(* PLC project boiler-plc210.project, CODESYS CODESYS V3.5 SP17 Patch 3 *)
(* stored: creationDateTime 2026-10-20T00:00:00, modificationDateTime 2026-10-20T00:00:00 *)
(* Синтетический экспорт: логика — corpus/boiler-plc210/src, слой ОВЕН — tools/corpus/owen_overlay.py (проба P7 не выполнялась) *)

// Назначение: состояние котла (вымышленная котельная №3, ПЛК210 — синтетический слой ОВЕН).
// Автор:      kr0nsch
// Версия:     0.1.0
// Документ:   corpus/boiler-plc210/README.md
{attribute 'qualified_only'}
TYPE E_BoilerState :
(
    Off := 0,       // остановлен
    Run := 1,       // работа
    Fault := 2      // авария горелки
) INT;
END_TYPE

// Назначение: отопительный график: уставка подачи по наружной температуре (линейно, с ограничением).
// Автор:      kr0nsch
// Версия:     0.1.0
// Документ:   corpus/boiler-plc210/README.md
FUNCTION F_HeatingCurve : REAL
VAR_INPUT
    rTOutdoor_C : REAL;     // наружная температура, °C
    rSpBase_C : REAL;       // уставка при 0 °C
END_VAR
VAR CONSTANT
    SLOPE : REAL := -1.2;   // наклон графика, °C/°C
    SP_MIN : REAL := 35.0;  // минимум подачи, °C
    SP_MAX : REAL := 95.0;  // максимум подачи, °C
END_VAR

            F_HeatingCurve := LIMIT(SP_MIN, rSpBase_C + SLOPE * rTOutdoor_C, SP_MAX);

          
END_FUNCTION

// Назначение: резервный электрокотёл — двухпозиционный регулятор ON_OFF_HIST_REG (CmpOwenPidRegs).
// Автор:      kr0nsch
// Версия:     0.1.0
// Документ:   corpus/boiler-plc210/README.md
PROGRAM PRG_Backup
VAR
    fbHeater : OPR.ON_OFF_HIST_REG; // двухпозиционный регулятор
    xHeaterOn : BOOL;               // включить ТЭН
END_VAR
VAR CONSTANT
    SP_BACKUP_C : REAL := 45.0;     // уставка резерва, °C
    HYST_C : REAL := 2.0;           // гистерезис, °C
END_VAR

            fbHeater(PV := GVL_Mx.rTSupply_C, SP := SP_BACKUP_C, HYST := HYST_C, DB := 0.0);
xHeaterOn := fbHeater.HEATER AND GVL_Hmi.eState = E_BoilerState.Fault;

          
END_PROGRAM

// Назначение: быстрые блокировки (задача FastTask, приоритет 0 у ОВЕН): авария горелки -> останов, сирена.
// Автор:      kr0nsch
// Версия:     0.1.0
// Документ:   corpus/boiler-plc210/README.md
PROGRAM PRG_Fast
VAR
END_VAR

            IF GVL_Hw.xBurner1Fault OR GVL_Hw.xBurner2Fault THEN
    GVL_Hmi.eState := E_BoilerState.Fault;
    GVL_Hw.xAlarmHorn := TRUE;
ELSE
    GVL_Hw.xAlarmHorn := FALSE;
END_IF

          
END_PROGRAM

// Назначение: регулирование подачи (ПИД CmpOwenPidRegs), насос, строки для панели (OwenStringUtils).
// Автор:      kr0nsch
// Версия:     0.1.0
// Документ:   corpus/boiler-plc210/README.md
PROGRAM PRG_Main
VAR
    fbPid : OPR.STD_PID;    // ПИД подачи
    rSp_C : REAL;           // уставка подачи, °C
    rValve : REAL;          // выход ПИД 0..1
    fbRunTimer : TON;       // секундный такт наработки
END_VAR
VAR CONSTANT
    XP_C : REAL := 20.0;    // полоса пропорциональности, °C
    TI_S : REAL := 120.0;   // постоянная интегрирования, с
    T_SECOND : TIME := T#1S;    // такт счёта наработки
    DIGITS : USINT := 1;    // знаков после запятой
END_VAR

            rSp_C := F_HeatingCurve(GVL_Mx.rTOutdoor_C, GVL_Persist.rSpBase_C);
fbPid(PV := GVL_Mx.rTSupply_C, SP := rSp_C, XP := XP_C, TI := TI_S, TD := 0.0, PMIN := 0.0, PMAX := 1.0,
      Y_MAN_SET := FALSE, Y_MANUAL := 0.0);
rValve := fbPid.Y;
IF GVL_Hmi.eState <> E_BoilerState.Fault THEN
    GVL_Hmi.eState := E_BoilerState.Run;
END_IF
GVL_Hw.xPumpRun := GVL_Hmi.eState = E_BoilerState.Run;
GVL_Mx.wDoMask := SEL(GVL_Hw.xPumpRun, 16#0000, 16#0001);
fbRunTimer(IN := GVL_Hw.xPumpRun AND NOT fbRunTimer.Q, PT := T_SECOND);
IF fbRunTimer.Q THEN
    GVL_Persist.udiRunTime_s := GVL_Persist.udiRunTime_s + 1;
END_IF
GVL_Hmi.sStatus := OSU.CONCAT4('T=', OSU.REAL_TO_STRING_FORMAT(GVL_Mx.rTSupply_C, DIGITS, OSU.DECIMAL_SEPARATOR.COMMA),
                               ' C, SP=', OSU.REAL_TO_STRING_FORMAT(rSp_C, DIGITS, OSU.DECIMAL_SEPARATOR.COMMA));
GVL_Hmi.sCode := OSU.WORD_TO_HEX_STR(wInput := GVL_Hw.wHmiStatus, xUpperCase := TRUE, sPrefix := '0x');

          
END_PROGRAM

// Назначение: медленная задача (приоритет 15 у ОВЕН): слово состояния панели.
// Автор:      kr0nsch
// Версия:     0.1.0
// Документ:   corpus/boiler-plc210/README.md
PROGRAM PRG_Slow
VAR
END_VAR
VAR CONSTANT
    BIT_FAULT : WORD := 16#0002;    // бит «авария» в слове состояния
    BIT_RUN : WORD := 16#0001;      // бит «работа»
END_VAR

            GVL_Hw.wHmiStatus := 0;
IF GVL_Hmi.eState = E_BoilerState.Run THEN
    GVL_Hw.wHmiStatus := GVL_Hw.wHmiStatus OR BIT_RUN;
END_IF
IF GVL_Hmi.eState = E_BoilerState.Fault THEN
    GVL_Hw.wHmiStatus := GVL_Hw.wHmiStatus OR BIT_FAULT;
END_IF

          
END_PROGRAM

CONFIGURATION Device
  RESOURCE Application ON PLC
(* global variable list GVL_Clock *)
// Назначение: время ПЛК из каналов узла OwenRTC и данные узла Watchdog.
// Автор:      kr0nsch
// Версия:     0.1.0
// Документ:   corpus/boiler-plc210/README.md
VAR_GLOBAL
    dtNow : DT;             // Date And Time
    sDateText : STRING(80); // Format date
    sTimeText : STRING(80); // Format time
    usiHour : USINT;        // Hour
    usiWeek : USINT;        // Week of year
    udiLastExc : UDINT;     // Watchdog: код последнего исключения
END_VAR
(* global variable list GVL_Hmi *)
// Назначение: строки и коды для панели оператора.
// Автор:      kr0nsch
// Версия:     0.1.0
// Документ:   corpus/boiler-plc210/README.md
VAR_GLOBAL
    sStatus : STRING(255);  // строка состояния
    sCode : STRING(8);      // код состояния (hex)
    eState : E_BoilerState; // состояние котла К1
END_VAR
(* global variable list GVL_Hw *)
// Назначение: встроенный ввод-вывод ПЛК210 по AT-адресам (так делать ОВЕН не рекомендует — Targets v3.4, разд. 1;
//             вход нарочно с AT, чтобы показать C2A-IO001).
// Автор:      kr0nsch
// Версия:     0.1.0
// Документ:   corpus/boiler-plc210/README.md
VAR_GLOBAL
    xBurner1Fault AT %IX0.0 : BOOL;     // авария горелки К1
    xBurner2Fault AT %IX0.1 : BOOL;     // авария горелки К2
    xPumpRun AT %QX0.0 : BOOL;          // пуск сетевого насоса Н1
    xAlarmHorn AT %QX0.1 : BOOL;        // сирена
    wHmiStatus AT %MW10 : WORD;         // слово состояния для панели
END_VAR
(* global variable list GVL_Mx *)
// Назначение: значения модулей Mx210 (привязки к каналам шаблонов МВ210-101 и МУ210-402 в дереве устройств).
// Автор:      kr0nsch
// Версия:     0.1.0
// Документ:   corpus/boiler-plc210/README.md
VAR_GLOBAL
    rTSupply_C : REAL;      // температура подачи, °C (МВ210-101, вход 1)
    rTReturn_C : REAL;      // температура обратки, °C (вход 2)
    rTOutdoor_C : REAL;     // температура наружного воздуха, °C (вход 3)
    iTSupplyRaw : INT;      // подача, целое (вход 1, integer)
    wDoMask : WORD;         // выходы МУ210-402 (битовая маска)
    wMeterStatus : WORD;    // счётчик энергии на Modbus 3S (канал FC 23)
END_VAR
(* global variable list GVL_Persist *)
// Назначение: сохраняемые уставки и наработка.
// Автор:      kr0nsch
// Версия:     0.1.0
// Документ:   corpus/boiler-plc210/README.md
VAR_GLOBAL RETAIN
    rSpBase_C : REAL := 70.0;   // базовая уставка подачи, °C
    udiRunTime_s : UDINT;       // наработка насоса, с
END_VAR
    TASK FastTask(INTERVAL := T#50ms, PRIORITY := 0);
    TASK MainTask(INTERVAL := T#50ms, PRIORITY := 1);
    TASK SlowTask(INTERVAL := T#50ms, PRIORITY := 15);
    PROGRAM PRG_Fast WITH FastTask : PRG_Fast;
    PROGRAM PRG_Main WITH MainTask : PRG_Main;
    PROGRAM PRG_Backup WITH MainTask : PRG_Backup;
    PROGRAM PRG_Slow WITH SlowTask : PRG_Slow;
  END_RESOURCE
END_CONFIGURATION

CONFIGURATION OwenRTC
END_CONFIGURATION

CONFIGURATION Watchdog
END_CONFIGURATION

CONFIGURATION Modbus_TCP_Master
END_CONFIGURATION

CONFIGURATION MV210_101_K3
END_CONFIGURATION

CONFIGURATION MU210_402_K3
END_CONFIGURATION

CONFIGURATION ModbusTCP_Slave_Device_Meter
END_CONFIGURATION
